(* IEC 61131-3 sources: tsplc/packages/vscode-extension/tests/fixtures/blueprint, 1 file *)

(* ---- Main.st ---- *)
PROGRAM Main
VAR
	Inbound : FB_ZoneConveyor;
END_VAR

(* Bind the conveyor each cycle before calling Inbound.SetMotionSignal(). *)
Inbound(Conveyor := PlantIO.Conveyor_Infeed);

END_PROGRAM
